Fanuc KAREL source: KT00174.KL

PROGRAM KT00174
%NOLOCKGROUP
VAR
  R1: REAL
  Y2: ARRAY[2] OF BYTE
  OUT: REAL
BEGIN
  R1 = 2.0
    Y2[1] = 3
  OUT = R1 MOD Y2[1]
END KT00174
